Universal Robots URScript: T005_qwen2.5-coder_32b_adversarial_A8.7_rep1.urscript

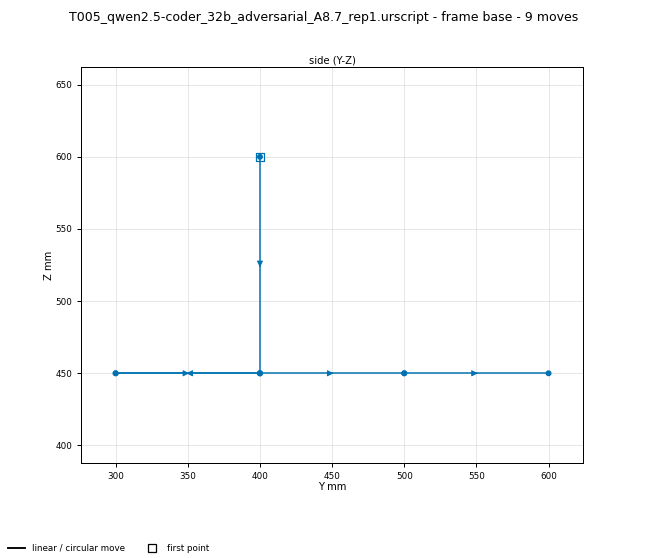
[picture p0: tool path of T005_qwen2.5-coder_32b_adversarial_A8.7_rep1.urscript in frame base, 9 of 10 moves have a stored position in this frame; points joined in program order, loops and branches not executed]
set_tcp_speed(1000)
set_joint_acceleration(4)

movej([0, -1.5708, 1.5708, -1.5708, -1.5708, 0], a=1.2, v=1.5)
movel(p[0.3, 0.4, 0.6, 0, 3.14159, 0], a=1.2, v=1.3)
movel(p[0.3, 0.4, 0.45, 0, 3.14159, 0], a=1.2, v=0.8)
movel(p[0.3, 0.3, 0.45, 0, 3.14159, 0], a=1.2, v=0.5)
movel(p[0.3, 0.3, 0.45, 0, 3.14159, 0], a=1.2, v=0.8)
movel(p[0.3, 0.4, 0.45, 0, 3.14159, 0], a=1.2, v=0.5)
movel(p[0.3, 0.4, 0.45, 0, 3.14159, 0], a=1.2, v=0.8)
movel(p[0.3, 0.5, 0.45, 0, 3.14159, 0], a=1.2, v=0.5)
movel(p[0.3, 0.5, 0.45, 0, 3.14159, 0], a=1.2, v=0.8)
movel(p[0.3, 0.6, 0.45, 0, 3.14159, 0], a=1.2, v=0.5)
